// TwinCAT 3 PLC project PLC1
// ProgramVersion: 3.1.4026.22
// CompilerDefines: VISU_USEPROPERTYINFO,VISU_USEWSTRING
// libraries:
//   Tc2_Standard, * (Beckhoff Automation GmbH)
//   Tc2_System, * (Beckhoff Automation GmbH)
//   VisuDialogs, * (System)
//   VisuSymbols, 4.5.0.0 (System)
// project tree:
//   / GlobalTextList.TcGTLO, PlcTask.TcTTO, VISU_TASK.TcTTO
//   GVLs/ GVL.TcGVL
//   POUs/ MAIN.TcPOU
//   VISUs/ Main.TcVIS, Visualization Manager.TcVMO (not stored)
// real-time tasks:
//   TASK PlcTask: cycle T#10ms, priority 20, ADS port 350
//   TASK VISU_TASK: cycle T#200000us, priority 30, ADS port 351

CONFIGURATION PLC1
    RESOURCE PLC ON TwinCAT3
        TASK PlcTask(INTERVAL := T#10ms, PRIORITY := 20);
        TASK VISU_TASK(INTERVAL := T#200000us, PRIORITY := 30);
        PROGRAM MAIN WITH PlcTask : MAIN;
        PROGRAM VisuElems_Visu_Prg WITH VISU_TASK : VisuElems.Visu_Prg;
    END_RESOURCE
END_CONFIGURATION

// ---- GVLs/GVL.TcGVL
{attribute 'qualified_only'}
VAR_GLOBAL
	    // =====================================================================
    // 場景 1:輸送帶分料站 — 與模擬器的介面
    //
    // PLC → 模擬器:致動器命令(由 PLC 程式寫入)
    // 模擬器 → PLC:感測器回饋(由模擬器寫入,PLC 只能讀)
    //
    // 注意:標示為「模擬器寫入」的變數請勿在 PLC 程式中賦值,
    //       否則每個週期都會被模擬器覆蓋,行為會很難除錯。
    // =====================================================================

    // ---------- PLC → 模擬器(致動器)----------
    bFeederRun          : BOOL;     // 進料機構啟動
    bBeltForward        : BOOL;     // 輸送帶正轉(往出料端)
    bBeltReverse        : BOOL;     // 輸送帶反轉(往進料端)
    bCylExtend          : BOOL;     // 氣缸推出電磁閥(單動,FALSE 自動縮回)
    bResetCounters      : BOOL;     // 計數歸零(持續為 TRUE 期間持續歸零)

    // ---------- 模擬器 → PLC(感測器)----------
    bSensorEntry        : BOOL;     // 進料感測器
    bSensorInspect      : BOOL;     // 檢測位感測器
    bSensorExit         : BOOL;     // 出料感測器
    bPartIsNg           : BOOL;     // 檢測位上的零件為 NG 品
    bCylExtended        : BOOL;     // 氣缸前限位
    bCylRetracted       : BOOL;     // 氣缸後限位
    bBeltFault          : BOOL;     // 正反轉同時給命令 → 皮帶停止並報異常
    rBeltPos            : LREAL;    // 皮帶累積位移 [mm](反轉時會減少)
    // 兩個都是「位置計數器」,不看零件好壞:
    // 分料沒推成功的 NG 品會計進 iCountOk,推錯的 OK 品會計進 iCountNg。
    // 拿它們跟實際投料比對,就能驗證分料邏輯寫得對不對。
    iCountOk            : DINT;     // 從出料端離開的總數
    iCountNg            : DINT;     // 被推入退料槽的總數
    iCountReturned      : DINT;     // 反轉退回進料端而流失的數量
	
	//HMI buttons
	bStart : BOOL;
	bStop  : BOOL;
	

END_VAR

// ---- POUs/MAIN.TcPOU
PROGRAM MAIN
VAR
	fbCTU1 : CTU;
	fbCTU2 : CTU;
	fbCTU3 : CTU;
	iState : INT;
	fbRtrigS1 : R_TRIG;
	fbRtrigS2 : R_TRIG;
	fbRtrigS3 : R_TRIG;
	
	
	
END_VAR

fbRtrigS1(CLK:=GVL.bSensorEntry , Q=> );
fbRtrigS2(CLK:=GVL.bSensorInspect , Q=> );
fbRtrigS3(CLK:=GVL.bSensorExit , Q=> );

fbCTU1(
	CU:= fbRtrigS1.Q , 
	RESET:= , 
	PV:=999 , 
	Q=> , 
	CV=> );
fbCTU2(CU:=fbRtrigS2.Q, PV:=999);
fbCTU3(CU:=fbRtrigS3.Q, PV:=999);

IF GVL.bStop THEN
	iState := 999;
END_IF


CASE iState OF 
	0:
		fbCTU1.RESET := TRUE;
		fbCTU2.RESET := TRUE;
		fbCTU3.RESET := TRUE;
		GVL.bBeltForward := FALSE;
		GVL.bBeltReverse := FALSE;		
		GVL.bCylExtend := FALSE;
		GVL.bFeederRun := FALSE;
		IF GVL.bStart THEN
			iState :=100;
		END_IF
		
	100:
		fbCTU1.RESET := FALSE;
		fbCTU2.RESET := FALSE;
		fbCTU3.RESET := FALSE;		
		GVL.bFeederRun := TRUE;
		GVL.bBeltForward := TRUE;
		IF GVL.bPartIsNg AND GVL.bSensorInspect THEN
			GVL.bCylExtend := TRUE;
		ELSIF GVL.bCylExtended THEN
			GVL.bCylExtend := FALSE; 
			
		END_IF
		IF fbCTU3.CV >=20 THEN
			iState :=200;
		END_IF
	200:
		GVL.bBeltForward := FALSE;
		GVL.bBeltReverse := FALSE;		
		GVL.bCylExtend := FALSE;
		GVL.bFeederRun := FALSE;
		iState :=0;
	999:
		GVL.bBeltForward := FALSE;
		GVL.bBeltReverse := FALSE;		
		GVL.bCylExtend := FALSE;
		GVL.bFeederRun := FALSE;
		IF GVL.bStart THEN
			iState :=100;
		END_IF

END_CASE

END_PROGRAM

// ---- GlobalTextList.TcGTLO
TEXTLIST GlobalTextList
  90 = '%s'
  239 = 'Start'
  245 = 'Stop'
END_TEXTLIST

// ---- VISUs/Main.TcVIS
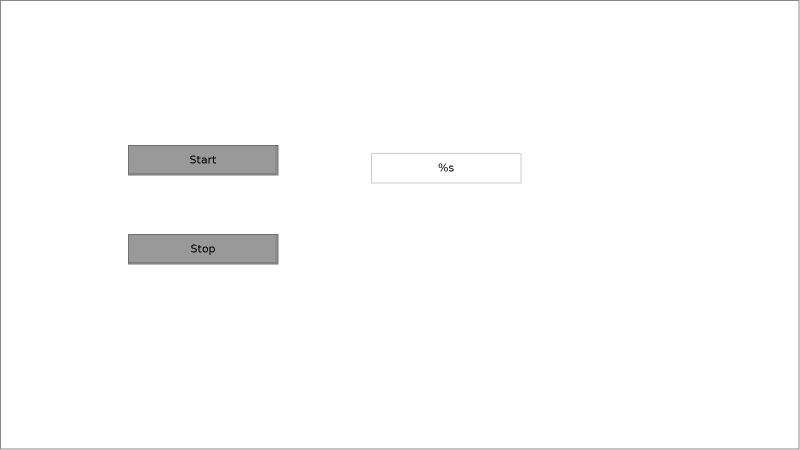
VISUALIZATION Main  // 800x450
    Button (128,145 150x30), "Start"
        tap GVL.bStart
    Button (128,234 150x30), "Stop"
        tap GVL.bStop
    Textfield (371,153 150x30), "%s", text variable: MAIN.fbCTU3.CV
END_VISUALIZATION
